TYPE ST_KUKA_REF_1 : FB_KUKA_REF;
END_TYPE

(* stored: Version 1.1.0.1, ProductVersion 3.1.4024.15
   DUT ST_KUKA_REF_1: Id {bddd25dc-b27a-4a38-9360-3e194961f293} *)
